(* IEC 61131-3 sources: repolevel_ST_code_completion/dataset/project_code/ProductionLine/struct, 2 files *)

(* ---- MotorI.st ---- *)
TYPE MotorI :
STRUCT
	Start:BOOL;
	Stop:BOOL;
	Overload:BOOL;
	FaultReset:BOOL;
END_STRUCT
END_TYPE

(* ---- MotorO.st ---- *)
TYPE MotorO :
STRUCT
	Coil:BOOL;
	FaultStatus:BOOL;
END_STRUCT
END_TYPE
